(* IEC 61131-3 sources: kns-pump-station/tests/POUs/Log/FB_AlarmSummary_Test, 18 files *)

(* ---- AckByIdDeviceStationPid.method.decl.st ---- *)
// Квитирование по номеру у источников с номерами устройства (110), станции (100005) и LIC101 (100100);
// чужой номер и повторное квитирование — FALSE
METHOD PRIVATE AckByIdDeviceStationPid
VAR_INST
    fbDut  : FB_AlarmSummary;       // проверяемая сводка
    stView : ST_AlarmView;          // список тревог
    fbDev  : FB_TestAlarmSource;    // «устройство»: тревоги 110, 111
    fbStn  : FB_TestAlarmSource;    // «станция»: тревога 100005
    fbPid  : FB_TestAlarmSource;    // «LIC101»: тревога 100100
END_VAR
VAR
    fbTime : PL.FB_FakeTime;        // подменное время
    itfAlm : PL.I_Alarm;            // проверяемая тревога источника
END_VAR

(* ---- CountsByPriority.method.decl.st ---- *)
// Активные Low, Medium, High неквитированные и Critical квитированная: активных по одной на приоритет,
// неквитированных — Low, Medium, High
METHOD PRIVATE CountsByPriority
VAR_INST
    fbDut  : FB_AlarmSummary;       // проверяемая сводка
    stView : ST_AlarmView;          // список тревог
    fbSrc1 : FB_TestAlarmSource;    // источник 1: Low, Medium, High
    fbSrc2 : FB_TestAlarmSource;    // источник 2: Critical
END_VAR
VAR
    fbTime : PL.FB_FakeTime;        // подменное время
END_VAR

(* ---- EmptyDefaults.method.decl.st ---- *)
// Без источников: счётчики 0, неквитированных нет, список пуст, первый вызов пересчитывает список
METHOD PRIVATE EmptyDefaults
VAR_INST
    fbDut  : FB_AlarmSummary;       // проверяемая сводка
    stView : ST_AlarmView;          // список тревог
END_VAR
VAR
    fbTime : PL.FB_FakeTime;        // подменное время
    uiI    : UINT;                  // приоритет
END_VAR

(* ---- EmptyDefaults.method.impl.st ---- *)
coUnit.TEST('AlarmSummary_EmptyDefaults');

fbDut(uiSourceCount := 0, itfTime := fbTime, stView := stView);
FOR uiI := 1 TO GVL_Const.ALM_PRIO_COUNT DO
    AssertEquals_UINT(Expected := 0, Actual := fbDut.auiActive[uiI] + fbDut.auiUnack[uiI], Message := 'counters 0');
END_FOR
AssertTrue(Condition := fbDut.ePrioUnack = PL.E_AlarmPriority.None, Message := 'no unacked');
AssertEquals_UINT(Expected := 0, Actual := stView.uiCount, Message := 'empty view');
AssertEquals_UDINT(Expected := 1, Actual := stView.udiRevision, Message := 'view built on first call');

coUnit.TEST_FINISHED();

(* ---- NewHighSeqOnlyOnTransition.method.decl.st ---- *)
// Счётчик новых High/Critical растёт только на переходе в ActiveUnack: держится, не растёт от Medium, снова
// растёт после возврата и повторного появления
METHOD PRIVATE NewHighSeqOnlyOnTransition
VAR_INST
    fbDut  : FB_AlarmSummary;       // проверяемая сводка
    stView : ST_AlarmView;          // список тревог
    fbSrc  : FB_TestAlarmSource;    // источник: High, Medium
END_VAR
VAR
    fbTime : PL.FB_FakeTime;        // подменное время
END_VAR

(* ---- PrioUnackHighest.method.decl.st ---- *)
// Высший неквитированный приоритет: Medium неквитирована, High квитирована → Medium; Critical появилась → Critical
METHOD PRIVATE PrioUnackHighest
VAR_INST
    fbDut  : FB_AlarmSummary;       // проверяемая сводка
    stView : ST_AlarmView;          // список тревог
    fbSrc  : FB_TestAlarmSource;    // источник: Medium, High, Critical
END_VAR
VAR
    fbTime : PL.FB_FakeTime;        // подменное время
END_VAR

(* ---- PrioUnackHighestBeforeLower.method.decl.st ---- *)
// Высший неквитированный приоритет не зависит от порядка обхода: Critical в слоте 0, Low в слоте 1 (обе
// неквитированы) → Critical, а не приоритет последней найденной
METHOD PRIVATE PrioUnackHighestBeforeLower
VAR_INST
    fbDut  : FB_AlarmSummary;       // проверяемая сводка
    stView : ST_AlarmView;          // список тревог
    fbSrc  : FB_TestAlarmSource;    // источник: Critical, Low
END_VAR
VAR
    fbTime : PL.FB_FakeTime;        // подменное время
END_VAR

(* ---- ShelveByIdRespectsTShelveMax.method.decl.st ---- *)
// Откладывание по номеру: tShelveMax = 0 — отказ; 1 ч — принято, через 1 ч откладывание истекает и активная
// тревога снова ActiveUnack
METHOD PRIVATE ShelveByIdRespectsTShelveMax
VAR_INST
    fbDut  : FB_AlarmSummary;       // проверяемая сводка
    stView : ST_AlarmView;          // список тревог
    fbSrc  : FB_TestAlarmSource;    // слот 0: откладывать нельзя; слот 1: до 1 ч
END_VAR
VAR
    fbTime : PL.FB_FakeTime;        // подменное время
    itfAlm : PL.I_Alarm;            // проверяемая тревога источника
END_VAR

(* ---- ShelveByIdUsesFullTShelveMax.method.decl.st ---- *)
// ShelveById откладывает на весь tShelveMax тревоги (по умолчанию 8 ч), а не на свой срок: через 1 ч 1 с тревога
// ещё отложена, через 8 ч 1 с — снова ActiveUnack
METHOD PRIVATE ShelveByIdUsesFullTShelveMax
VAR_INST
    fbDut  : FB_AlarmSummary;       // проверяемая сводка
    stView : ST_AlarmView;          // список тревог
    fbSrc  : FB_TestAlarmSource;    // слот 0: tShelveMax по умолчанию (8 ч)
END_VAR
VAR
    fbTime : PL.FB_FakeTime;        // подменное время
    itfAlm : PL.I_Alarm;            // проверяемая тревога источника
END_VAR

(* ---- StationSlotsBeyondDeviceLimit.method.decl.st ---- *)
// PMI-01, PMI-30: у станции 13 тревог (slot 1…13), у устройства библиотеки — до восьми. Сводка видит все слоты
// источника: KNS1.SIM (slot 13) и KNS1.NOAUTO (slot 9) попадают в счётчики, в список тревог и квитируются по номеру
METHOD PRIVATE StationSlotsBeyondDeviceLimit
VAR_INST
    fbDut  : FB_AlarmSummary;       // проверяемая сводка
    stView : ST_AlarmView;          // список тревог
    fbStn  : FB_StationAlarms;      // настоящий источник станции: 13 тревог
    stCfg  : ST_StationCfg;         // тревоги станции по умолчанию (05_alarm_list.csv)
END_VAR
VAR
    fbTime : PL.FB_FakeTime;        // подменное время
    itfAlm : PL.I_Alarm;            // проверяемая тревога источника
END_VAR

(* ---- TimeBackwardsRebuildsView.method.decl.st ---- *)
// «Время назад»: список пересчитывается сразу (разность LTIME без знака не считается)
METHOD PRIVATE TimeBackwardsRebuildsView
VAR_INST
    fbDut  : FB_AlarmSummary;       // проверяемая сводка
    stView : ST_AlarmView;          // список тревог
END_VAR
VAR
    fbTime : PL.FB_FakeTime;        // подменное время
END_VAR

(* ---- UnshelveById.method.decl.st ---- *)
// Возврат отложенной тревоги по номеру: TRUE и снова ActiveUnack; повторно — FALSE (не отложена)
METHOD PRIVATE UnshelveById
VAR_INST
    fbDut  : FB_AlarmSummary;       // проверяемая сводка
    stView : ST_AlarmView;          // список тревог
    fbSrc  : FB_TestAlarmSource;    // одна тревога
END_VAR
VAR
    fbTime : PL.FB_FakeTime;        // подменное время
    itfAlm : PL.I_Alarm;            // проверяемая тревога источника
END_VAR

(* ---- ViewLimitedToRows.method.decl.st ---- *)
// 56 активных тревог (7 источников по 8): в списке ALM_VIEW_ROWS строк, uiActiveTotal — настоящее число
METHOD PRIVATE ViewLimitedToRows
VAR_INST
    fbDut  : FB_AlarmSummary;       // проверяемая сводка
    stView : ST_AlarmView;          // список тревог
    afbSrc : ARRAY[1..7] OF FB_TestAlarmSource;   // источники по 8 тревог
END_VAR
VAR
    fbTime : PL.FB_FakeTime;        // подменное время
    uiS    : UINT;                  // источник
    uiK    : UINT;                  // слот
END_VAR

(* ---- ViewLimitedToRows.method.impl.st ---- *)
coUnit.TEST('AlarmSummary_ViewLimitedToRows');

FOR uiS := 1 TO 7 DO
    FOR uiK := 0 TO GVL_Const.ALM_SLOT_MAX DO
        afbSrc[uiS].axIn[uiK] := TRUE;
    END_FOR
    afbSrc[uiS](uiSlots := GVL_Const.ALM_SLOT_MAX + 1, udiIdBase := uiS * 100, itfTime := fbTime);
    fbDut.aitfSource[uiS] := afbSrc[uiS];
END_FOR
fbDut(uiSourceCount := 7, itfTime := fbTime, stView := stView);
AssertEquals_UINT(Expected := GVL_Const.ALM_VIEW_ROWS, Actual := stView.uiCount, Message := 'view limited to 50');
AssertEquals_UINT(Expected := 56, Actual := stView.uiActiveTotal, Message := 'total 56');
AssertEquals_UINT(Expected := 56, Actual := fbDut.auiUnack[2], Message := '56 unacked Medium');
AssertTrue(Condition := stView.astRow[GVL_Const.ALM_VIEW_ROWS].udiId <> 0, Message := 'last row filled');

coUnit.TEST_FINISHED();

(* ---- ViewNewerFirstInGroup.method.decl.st ---- *)
// Внутри группы и приоритета новые выше: три неквитированные Medium, появившиеся с интервалом 1 с (№ 150, 151,
// 152), — в списке 152, 151, 150
METHOD PRIVATE ViewNewerFirstInGroup
VAR_INST
    fbDut  : FB_AlarmSummary;       // проверяемая сводка
    stView : ST_AlarmView;          // список тревог
    fbSrc  : FB_TestAlarmSource;    // слоты 0…2, Medium
END_VAR
VAR
    fbTime : PL.FB_FakeTime;        // подменное время
    uiK    : UINT;                  // слот
END_VAR

(* ---- ViewNewerFirstInGroup.method.impl.st ---- *)
coUnit.TEST('AlarmSummary_ViewNewerFirstInGroup');

fbDut.aitfSource[1] := fbSrc;
fbSrc(uiSlots := 3, udiIdBase := 150, itfTime := fbTime);
fbDut(uiSourceCount := 1, itfTime := fbTime, stView := stView);
FOR uiK := 0 TO 2 DO
    fbTime.Advance(tStep := T#1S);
    fbSrc.axIn[uiK] := TRUE;
    fbSrc(itfTime := fbTime);
    fbDut(itfTime := fbTime, stView := stView);
END_FOR
fbTime.Advance(tStep := GVL_Const.ALM_VIEW_PERIOD);
fbDut(itfTime := fbTime, stView := stView);
AssertEquals_UINT(Expected := 3, Actual := stView.uiCount, Message := '3 rows');
AssertEquals_UDINT(Expected := 152, Actual := stView.astRow[1].udiId, Message := 'newest first');
AssertEquals_UDINT(Expected := 151, Actual := stView.astRow[2].udiId, Message := 'middle');
AssertEquals_UDINT(Expected := 150, Actual := stView.astRow[3].udiId, Message := 'oldest last');

coUnit.TEST_FINISHED();

(* ---- ViewPeriodRespected.method.decl.st ---- *)
// Список пересчитывается раз в ALM_VIEW_PERIOD (500 мс): через 100 мс — нет, через 500 мс — да
METHOD PRIVATE ViewPeriodRespected
VAR_INST
    fbDut  : FB_AlarmSummary;       // проверяемая сводка
    stView : ST_AlarmView;          // список тревог
    fbSrc  : FB_TestAlarmSource;    // источник с одной тревогой
END_VAR
VAR
    fbTime : PL.FB_FakeTime;        // подменное время
END_VAR

(* ---- ViewSortedUnackFirst.method.decl.st ---- *)
// Порядок списка: неквитированные (Medium выше Low), затем активные квитированные (High), затем отложенные
METHOD PRIVATE ViewSortedUnackFirst
VAR_INST
    fbDut  : FB_AlarmSummary;       // проверяемая сводка
    stView : ST_AlarmView;          // список тревог
    fbSrc  : FB_TestAlarmSource;    // слоты: 0 Low, 1 High (квитирована), 2 Medium, 3 Medium (отложена)
END_VAR
VAR
    fbTime : PL.FB_FakeTime;        // подменное время
END_VAR
